SUBAPPLICATION logiBUS_AI_Calibrate_3P_IDA_Param_OPC (* logiBUS_AI_IDA (Analog-Eingang) mit 3-Punkt-Kalibrierung (AR_CALIBRATE_3P_REF, unabhaengig gespeicherte Rohwerte X_MIN/X_MID/X_MAX + Referenzwerte MIN_REF/MID_REF/MAX_REF alle INI-persistiert) auf VT-Zahlenfelder (Rohwert + kalibrierter Wert, je eigene CNumberVariable) + Bargraph (kalibriert) + 3 VT-Tasten (C_MIN/C_MID/C_MAX) + OPC-UA (Rohwert DWORD + kalibrierter Wert REAL, generisch, ein Kanal). Fuer Sensoren mit definierter Mittelstellung (z.B. Lenkwinkelsensor: links/geradeaus/rechts) statt reiner 2-Punkt-Linearisierung. *)
  (* Standard: 61499-2; Description: Copyright (c) 2026 Meisterschulen am Ostbahnhof This program and the accompanying materials are made available under the terms of the Eclipse Public License 2.0 which is available at https://www.eclipse.org/legal/epl-2.0/ SPDX-License-Identifier: EPL-2.0 *)
  (* Version 1.0, 2026-10-30, Franz Höpfinger, Meisterschulen am Ostbahnhof, Kopie von logiBUS_AI_Calibrate_3P_IDA_OPC (v1.12), InputRaw jetzt logiBUS_AI_Raw_VT_AR_Param_OPC: Hysterese/TimeDelta/TimeRateLimit des AI per Web + INI einstellbar (gleiche sSection). Zuerst fuer Achslenkung Winkel (pendelte beim Zentrieren). PublishCal auf AR_TO_Q_Publish_Fast_OPC: CAL-Publish (Self-Subscribe der Mittelpunkt-Automatik) ungedrosselt, nur VT-Anzeige 500 ms. *)
  PACKAGE MyLib::sys;
  IMPORT isobus::UT::Q::const::IDs::ID_NULL;
  IMPORT logiBUS::io::AI::logiBUS_AI;
  IMPORT logiBUS::io::AI::logiBUS_AI_S;
  IMPORT logiBUS::utils::conversion::phys::NumericObjectPool_S;
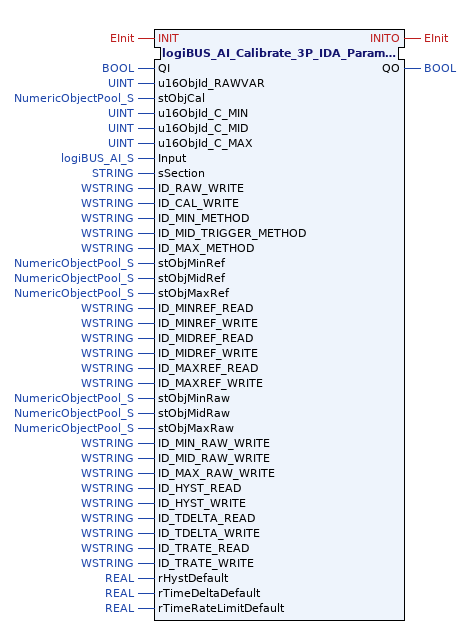
  EVENT_INPUT
    INIT : EInit; (* Initialization Request *)
  END_EVENT
  EVENT_OUTPUT
    INITO : EInit; (* Initialization Confirm *)
  END_EVENT
  VAR_INPUT
    QI : BOOL := TRUE; (* Quality Input - TRUE to enable service *)
    u16ObjId_RAWVAR : UINT := ID_NULL; (* Object ID CNumberVariable (Rohwert 0-4095, unkalibriert, reine Diagnose-Anzeige) *)
    stObjCal : logiBUS::utils::conversion::phys::NumericObjectPool_S := (u16ObjId := ID_NULL, r32Scale := 1.0, i32Offset := 0, u8Decimals := 1); (* Object ID + Scale/Offset/Decimals CNumberVariable (kalibrierter Wert, eigene, unabhaengige CNumberVariable) *)
    u16ObjId_C_MIN : UINT := ID_NULL; (* Object ID Taste 'C_MIN' (Min-Position anfahren, dann druecken) *)
    u16ObjId_C_MID : UINT := ID_NULL; (* Object ID Taste 'C_MID' (Mittelstellung anfahren, dann druecken) *)
    u16ObjId_C_MAX : UINT := ID_NULL; (* Object ID Taste 'C_MAX' (Max-Position anfahren, dann druecken) *)
    Input : logiBUS::io::AI::logiBUS_AI_S := logiBUS_AI::Invalid; (* Identify the Input AnalogInput_I1..I8 *)
    sSection : STRING; (* INI-Sektionsname fuer X_MIN/X_MID/X_MAX/MIN_REF/MID_REF/MAX_REF-Persistenz - pro Kanal eindeutig, sonst kollidieren die Kanaele in settings.ini *)
    ID_RAW_WRITE : WSTRING; (* Rohwert-Ruckmelde-Adresse (DWORD 0-4095, ACTION=PUBLISH) *)
    ID_CAL_WRITE : WSTRING; (* Kalibrierter-Wert-Ruckmelde-Adresse (REAL, ACTION=PUBLISH) *)
    ID_MIN_METHOD : WSTRING; (* Methodenadresse (ACTION=CREATE_METHOD) fuer den argumentlosen C_MIN-Trigger - gleichberechtigt zur lokalen VT-Taste aufrufbar, sowohl vom OPC-UA-Dashboard als auch per CLIENT_0 von einer anderen Station (siehe OPC_UA_VERNETZUNG.md Punkt 14 - kein Toggle/Subscribe-Umweg mehr) *)
    ID_MID_TRIGGER_METHOD : WSTRING; (* Methodenadresse (ACTION=CREATE_METHOD) fuer den argumentlosen C_MID-Trigger - siehe ID_MIN_METHOD *)
    ID_MAX_METHOD : WSTRING; (* Methodenadresse (ACTION=CREATE_METHOD) fuer den argumentlosen C_MAX-Trigger - siehe ID_MIN_METHOD *)
    stObjMinRef : logiBUS::utils::conversion::phys::NumericObjectPool_S := (u16ObjId := ID_NULL, r32Scale := 1.0, i32Offset := 0, u8Decimals := 1); (* Object ID + Scale/Offset/Decimals CNumberVariable (MIN_REF-Referenzwert, VT-Eingabefeld + OPC-UA) *)
    stObjMidRef : logiBUS::utils::conversion::phys::NumericObjectPool_S := (u16ObjId := ID_NULL, r32Scale := 1.0, i32Offset := 0, u8Decimals := 1); (* Object ID + Scale/Offset/Decimals CNumberVariable (MID_REF-Referenzwert, VT-Eingabefeld + OPC-UA) *)
    stObjMaxRef : logiBUS::utils::conversion::phys::NumericObjectPool_S := (u16ObjId := ID_NULL, r32Scale := 1.0, i32Offset := 0, u8Decimals := 1); (* Object ID + Scale/Offset/Decimals CNumberVariable (MAX_REF-Referenzwert, VT-Eingabefeld + OPC-UA) *)
    ID_MINREF_READ : WSTRING; (* Remote-Subscribe-Adresse MIN_REF-Referenzwert (REAL, ACTION=SUBSCRIBE) *)
    ID_MINREF_WRITE : WSTRING; (* Remote-Echo-Adresse MIN_REF-Referenzwert (REAL, ACTION=PUBLISH) *)
    ID_MIDREF_READ : WSTRING; (* Remote-Subscribe-Adresse MID_REF-Referenzwert (REAL, ACTION=SUBSCRIBE) *)
    ID_MIDREF_WRITE : WSTRING; (* Remote-Echo-Adresse MID_REF-Referenzwert (REAL, ACTION=PUBLISH) *)
    ID_MAXREF_READ : WSTRING; (* Remote-Subscribe-Adresse MAX_REF-Referenzwert (REAL, ACTION=SUBSCRIBE) *)
    ID_MAXREF_WRITE : WSTRING; (* Remote-Echo-Adresse MAX_REF-Referenzwert (REAL, ACTION=PUBLISH) *)
    stObjMinRaw : logiBUS::utils::conversion::phys::NumericObjectPool_S := (u16ObjId := ID_NULL, r32Scale := 1.0, i32Offset := 0, u8Decimals := 1); (* Object ID + Scale/Offset/Decimals CNumberVariable (Rohwert am MIN-Kalibrierpunkt, reine Diagnose-Anzeige) *)
    stObjMidRaw : logiBUS::utils::conversion::phys::NumericObjectPool_S := (u16ObjId := ID_NULL, r32Scale := 1.0, i32Offset := 0, u8Decimals := 1); (* Object ID + Scale/Offset/Decimals CNumberVariable (Rohwert am MID-Kalibrierpunkt, reine Diagnose-Anzeige) *)
    stObjMaxRaw : logiBUS::utils::conversion::phys::NumericObjectPool_S := (u16ObjId := ID_NULL, r32Scale := 1.0, i32Offset := 0, u8Decimals := 1); (* Object ID + Scale/Offset/Decimals CNumberVariable (Rohwert am MAX-Kalibrierpunkt, reine Diagnose-Anzeige) *)
    ID_MIN_RAW_WRITE : WSTRING; (* Rohwert-am-MIN-Kalibrierpunkt-Publish-Adresse (REAL, ACTION=PUBLISH) *)
    ID_MID_RAW_WRITE : WSTRING; (* Rohwert-am-MID-Kalibrierpunkt-Publish-Adresse (REAL, ACTION=PUBLISH) *)
    ID_MAX_RAW_WRITE : WSTRING; (* Rohwert-am-MAX-Kalibrierpunkt-Publish-Adresse (REAL, ACTION=PUBLISH) *)
    ID_HYST_READ : WSTRING; (* Web-Override AI-Hysterese (Digits) *)
    ID_HYST_WRITE : WSTRING; (* Rueckmeldung AI-Hysterese *)
    ID_TDELTA_READ : WSTRING; (* Web-Override AI-TimeDelta (ms) *)
    ID_TDELTA_WRITE : WSTRING; (* Rueckmeldung AI-TimeDelta *)
    ID_TRATE_READ : WSTRING; (* Web-Override AI-TimeRateLimit (ms) *)
    ID_TRATE_WRITE : WSTRING; (* Rueckmeldung AI-TimeRateLimit *)
    rHystDefault : REAL := 3.0; (* Default AI-Hysterese (Digits) *)
    rTimeDeltaDefault : REAL := 100.0; (* Default AI-TimeDelta (ms) *)
    rTimeRateLimitDefault : REAL := 20.0; (* Default AI-TimeRateLimit (ms) *)
  END_VAR
  VAR_OUTPUT
    QO : BOOL; (* Quality Output - TRUE if service executed successfully *)
  END_VAR
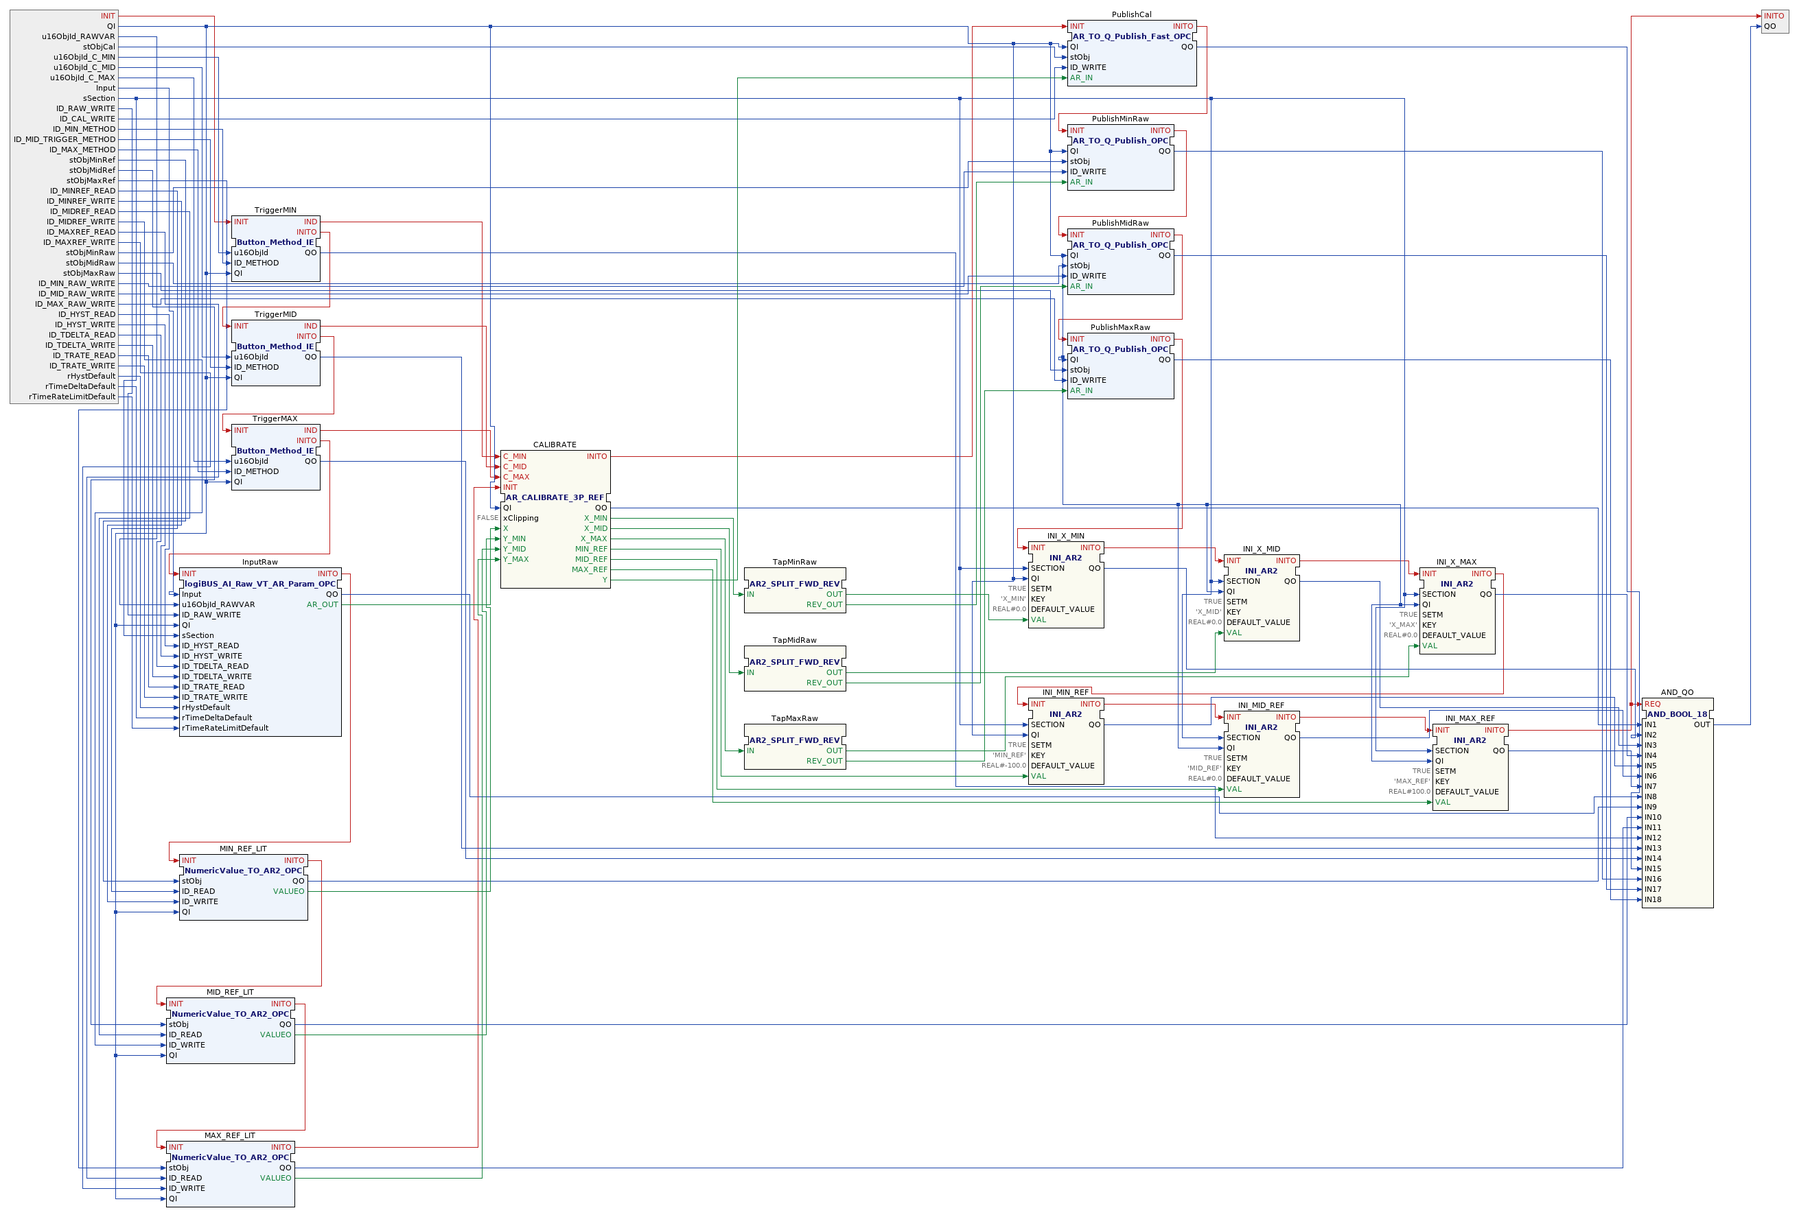
  FBS
    CALIBRATE : adapter::Engineering::measurements::AR_CALIBRATE_3P_REF(xClipping := FALSE);
    INI_X_MIN : eclipse4diac::storage::INI_AR2(SETM := TRUE, KEY := 'X_MIN', DEFAULT_VALUE := REAL#0.0);
    INI_X_MID : eclipse4diac::storage::INI_AR2(SETM := TRUE, KEY := 'X_MID', DEFAULT_VALUE := REAL#0.0);
    INI_X_MAX : eclipse4diac::storage::INI_AR2(SETM := TRUE, KEY := 'X_MAX', DEFAULT_VALUE := REAL#0.0);
    INI_MIN_REF : eclipse4diac::storage::INI_AR2(SETM := TRUE, KEY := 'MIN_REF', DEFAULT_VALUE := REAL#-100.0);
    INI_MID_REF : eclipse4diac::storage::INI_AR2(SETM := TRUE, KEY := 'MID_REF', DEFAULT_VALUE := REAL#0.0);
    INI_MAX_REF : eclipse4diac::storage::INI_AR2(SETM := TRUE, KEY := 'MAX_REF', DEFAULT_VALUE := REAL#100.0);
    TapMinRaw : adapter::events::bidirectional::AR2_SPLIT_FWD_REV;
    TapMidRaw : adapter::events::bidirectional::AR2_SPLIT_FWD_REV;
    TapMaxRaw : adapter::events::bidirectional::AR2_SPLIT_FWD_REV;
    AND_QO : iec61131::booleanOperators::AND_BOOL_18;
  END_FBS
  SUBAPPS
    InputRaw : MyLib::sys::logiBUS_AI_Raw_VT_AR_Param_OPC;
    MIN_REF_LIT : MyLib::sys::NumericValue_TO_AR2_OPC;
    MID_REF_LIT : MyLib::sys::NumericValue_TO_AR2_OPC;
    MAX_REF_LIT : MyLib::sys::NumericValue_TO_AR2_OPC;
    TriggerMIN : MyLib::sys::Button_Method_IE;
    TriggerMID : MyLib::sys::Button_Method_IE;
    TriggerMAX : MyLib::sys::Button_Method_IE;
    PublishCal : MyLib::sys::AR_TO_Q_Publish_Fast_OPC;
    PublishMinRaw : MyLib::sys::AR_TO_Q_Publish_OPC;
    PublishMidRaw : MyLib::sys::AR_TO_Q_Publish_OPC;
    PublishMaxRaw : MyLib::sys::AR_TO_Q_Publish_OPC;
  END_SUBAPPS
  EVENT_CONNECTIONS
    TriggerMIN.IND TO CALIBRATE.C_MIN;
    TriggerMID.IND TO CALIBRATE.C_MID;
    TriggerMAX.IND TO CALIBRATE.C_MAX;
    INIT TO TriggerMIN.INIT;
    CALIBRATE.INITO TO PublishCal.INIT;
    INI_X_MIN.INITO TO INI_X_MID.INIT;
    INI_X_MID.INITO TO INI_X_MAX.INIT;
    INI_X_MAX.INITO TO INI_MIN_REF.INIT;
    INI_MIN_REF.INITO TO INI_MID_REF.INIT;
    INI_MID_REF.INITO TO INI_MAX_REF.INIT;
    InputRaw.INITO TO MIN_REF_LIT.INIT;
    MIN_REF_LIT.INITO TO MID_REF_LIT.INIT;
    MID_REF_LIT.INITO TO MAX_REF_LIT.INIT;
    TriggerMIN.INITO TO TriggerMID.INIT;
    TriggerMID.INITO TO TriggerMAX.INIT;
    PublishCal.INITO TO PublishMinRaw.INIT;
    PublishMinRaw.INITO TO PublishMidRaw.INIT;
    PublishMidRaw.INITO TO PublishMaxRaw.INIT;
    INI_MAX_REF.INITO TO INITO;
    INI_MAX_REF.INITO TO AND_QO.REQ;
    TriggerMAX.INITO TO InputRaw.INIT;
    MAX_REF_LIT.INITO TO CALIBRATE.INIT;
    PublishMaxRaw.INITO TO INI_X_MIN.INIT;
  END_CONNECTIONS
  DATA_CONNECTIONS
    Input TO InputRaw.Input;
    u16ObjId_RAWVAR TO InputRaw.u16ObjId_RAWVAR;
    stObjCal TO PublishCal.stObj;
    u16ObjId_C_MIN TO TriggerMIN.u16ObjId;
    u16ObjId_C_MID TO TriggerMID.u16ObjId;
    u16ObjId_C_MAX TO TriggerMAX.u16ObjId;
    sSection TO INI_X_MIN.SECTION;
    sSection TO INI_X_MID.SECTION;
    sSection TO INI_X_MAX.SECTION;
    sSection TO INI_MIN_REF.SECTION;
    sSection TO INI_MID_REF.SECTION;
    sSection TO INI_MAX_REF.SECTION;
    ID_RAW_WRITE TO InputRaw.ID_RAW_WRITE;
    ID_CAL_WRITE TO PublishCal.ID_WRITE;
    ID_MIN_METHOD TO TriggerMIN.ID_METHOD;
    ID_MID_TRIGGER_METHOD TO TriggerMID.ID_METHOD;
    ID_MAX_METHOD TO TriggerMAX.ID_METHOD;
    stObjMinRef TO MIN_REF_LIT.stObj;
    ID_MINREF_READ TO MIN_REF_LIT.ID_READ;
    ID_MINREF_WRITE TO MIN_REF_LIT.ID_WRITE;
    stObjMidRef TO MID_REF_LIT.stObj;
    ID_MIDREF_READ TO MID_REF_LIT.ID_READ;
    ID_MIDREF_WRITE TO MID_REF_LIT.ID_WRITE;
    stObjMaxRef TO MAX_REF_LIT.stObj;
    ID_MAXREF_READ TO MAX_REF_LIT.ID_READ;
    ID_MAXREF_WRITE TO MAX_REF_LIT.ID_WRITE;
    stObjMinRaw TO PublishMinRaw.stObj;
    ID_MIN_RAW_WRITE TO PublishMinRaw.ID_WRITE;
    stObjMidRaw TO PublishMidRaw.stObj;
    ID_MID_RAW_WRITE TO PublishMidRaw.ID_WRITE;
    stObjMaxRaw TO PublishMaxRaw.stObj;
    ID_MAX_RAW_WRITE TO PublishMaxRaw.ID_WRITE;
    QI TO CALIBRATE.QI;
    QI TO INI_X_MIN.QI;
    QI TO INI_X_MID.QI;
    QI TO INI_X_MAX.QI;
    QI TO INI_MIN_REF.QI;
    QI TO INI_MID_REF.QI;
    QI TO INI_MAX_REF.QI;
    QI TO InputRaw.QI;
    QI TO MIN_REF_LIT.QI;
    QI TO MID_REF_LIT.QI;
    QI TO MAX_REF_LIT.QI;
    QI TO TriggerMIN.QI;
    QI TO TriggerMID.QI;
    QI TO TriggerMAX.QI;
    QI TO PublishCal.QI;
    QI TO PublishMinRaw.QI;
    QI TO PublishMidRaw.QI;
    QI TO PublishMaxRaw.QI;
    CALIBRATE.QO TO AND_QO.IN1;
    INI_X_MIN.QO TO AND_QO.IN2;
    INI_X_MID.QO TO AND_QO.IN3;
    INI_X_MAX.QO TO AND_QO.IN4;
    INI_MIN_REF.QO TO AND_QO.IN5;
    INI_MID_REF.QO TO AND_QO.IN6;
    INI_MAX_REF.QO TO AND_QO.IN7;
    InputRaw.QO TO AND_QO.IN8;
    MIN_REF_LIT.QO TO AND_QO.IN9;
    MID_REF_LIT.QO TO AND_QO.IN10;
    MAX_REF_LIT.QO TO AND_QO.IN11;
    TriggerMIN.QO TO AND_QO.IN12;
    TriggerMID.QO TO AND_QO.IN13;
    TriggerMAX.QO TO AND_QO.IN14;
    PublishCal.QO TO AND_QO.IN15;
    PublishMinRaw.QO TO AND_QO.IN16;
    PublishMidRaw.QO TO AND_QO.IN17;
    PublishMaxRaw.QO TO AND_QO.IN18;
    AND_QO.OUT TO QO;
    sSection TO InputRaw.sSection;
    ID_HYST_READ TO InputRaw.ID_HYST_READ;
    ID_HYST_WRITE TO InputRaw.ID_HYST_WRITE;
    ID_TDELTA_READ TO InputRaw.ID_TDELTA_READ;
    ID_TDELTA_WRITE TO InputRaw.ID_TDELTA_WRITE;
    ID_TRATE_READ TO InputRaw.ID_TRATE_READ;
    ID_TRATE_WRITE TO InputRaw.ID_TRATE_WRITE;
    rHystDefault TO InputRaw.rHystDefault;
    rTimeDeltaDefault TO InputRaw.rTimeDeltaDefault;
    rTimeRateLimitDefault TO InputRaw.rTimeRateLimitDefault;
  END_CONNECTIONS
  ADAPTER_CONNECTIONS
    InputRaw.AR_OUT TO CALIBRATE.X;
    CALIBRATE.X_MIN TO TapMinRaw.IN;
    TapMinRaw.OUT TO INI_X_MIN.VAL;
    TapMinRaw.REV_OUT TO PublishMinRaw.AR_IN;
    CALIBRATE.X_MID TO TapMidRaw.IN;
    TapMidRaw.OUT TO INI_X_MID.VAL;
    TapMidRaw.REV_OUT TO PublishMidRaw.AR_IN;
    CALIBRATE.X_MAX TO TapMaxRaw.IN;
    TapMaxRaw.OUT TO INI_X_MAX.VAL;
    TapMaxRaw.REV_OUT TO PublishMaxRaw.AR_IN;
    CALIBRATE.MIN_REF TO INI_MIN_REF.VAL;
    CALIBRATE.MID_REF TO INI_MID_REF.VAL;
    CALIBRATE.MAX_REF TO INI_MAX_REF.VAL;
    MIN_REF_LIT.VALUEO TO CALIBRATE.Y_MIN;
    MID_REF_LIT.VALUEO TO CALIBRATE.Y_MID;
    MAX_REF_LIT.VALUEO TO CALIBRATE.Y_MAX;
    CALIBRATE.Y TO PublishCal.AR_IN;
  END_CONNECTIONS
END_SUBAPPLICATION
